(* Logix 5000 project; controller CIP vendor 1 type 14 code 106 rev 20.12; software revision 20.06; part 3 of 13 *)
(* tags used below, declared in another part *)
   Alarm_Preset_Indx : DINT;
   Alarm_Timer : TIMER[128];
   Alarm_Timer_Preset : DINT[128];
   Bit : BOOL[128];
   Counter : COUNTER[10];
   Integer_1 : ALIAS FOR Integer[1];
   Integer_6 : ALIAS FOR Integer[6];
   One_Shot : BOOL[128];
   Panelview : INT[40];
   PV_Current_Select_Step_Op : DINT;
   PV_Edit_Opcodes : DINT[300];
   PV_Edit_Recipe_Name : STRING;
   PV_Edit_Recipe_Top_Row : DINT;
   PV_Edit_Recipes : DINT[7];
   PV_Edit_Recipes_0 : ALIAS FOR PV_Edit_Recipes[0];
   PV_Edit_Recipes_0_Prev : DINT;
   PV_Edit_Screen_Opcodes : DINT[17];
   PV_Edit_Setpoints : REAL[97];
   PV_Edit_Times : DINT[300];
   PV_Rename_Recipe_Name : STRING;
   PV_Security : Security_Main_HMI;
   PV_Security1 : Security_Remote_HMI;
   PV_Step_Time : REAL;
   PV_Visibility : INT[5];
   Recipe : RECIPE[41];
   Recipe_Name : STRING[41];
   Recipe_Name_Indx : DINT;
   SecurityLevel : DINT;
   SecurityLevel1 : DINT;
   Time_Date : DINT[20];
   WashChamberDoorGasketCTRL : DINT;
(* MainProgram, continued *)

ROUTINE _03_PV_SECURITY_REMOTE1_HMI   (* ladder *)
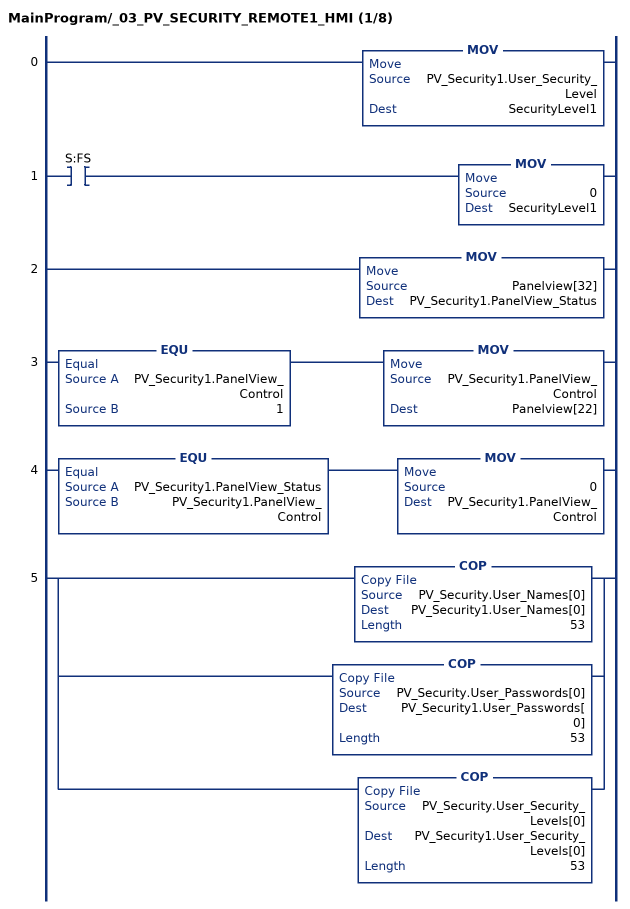
   0: MOV(PV_Security1.User_Security_Level,SecurityLevel1);
   1: XIC(S:FS)MOV(0,SecurityLevel1);
   2: MOV(Panelview[32],PV_Security1.PanelView_Status);
   3: EQU(PV_Security1.PanelView_Control,1)MOV(PV_Security1.PanelView_Control,Panelview[22]);
   4: EQU(PV_Security1.PanelView_Status,PV_Security1.PanelView_Control)MOV(0,PV_Security1.PanelView_Control);
   5: [COP(PV_Security.User_Names[0],PV_Security1.User_Names[0],53) ,COP(PV_Security.User_Passwords[0],PV_Security1.User_Passwords[0],53) ,COP(PV_Security.User_Security_Levels[0],PV_Security1.User_Security_Levels[0],53) ];
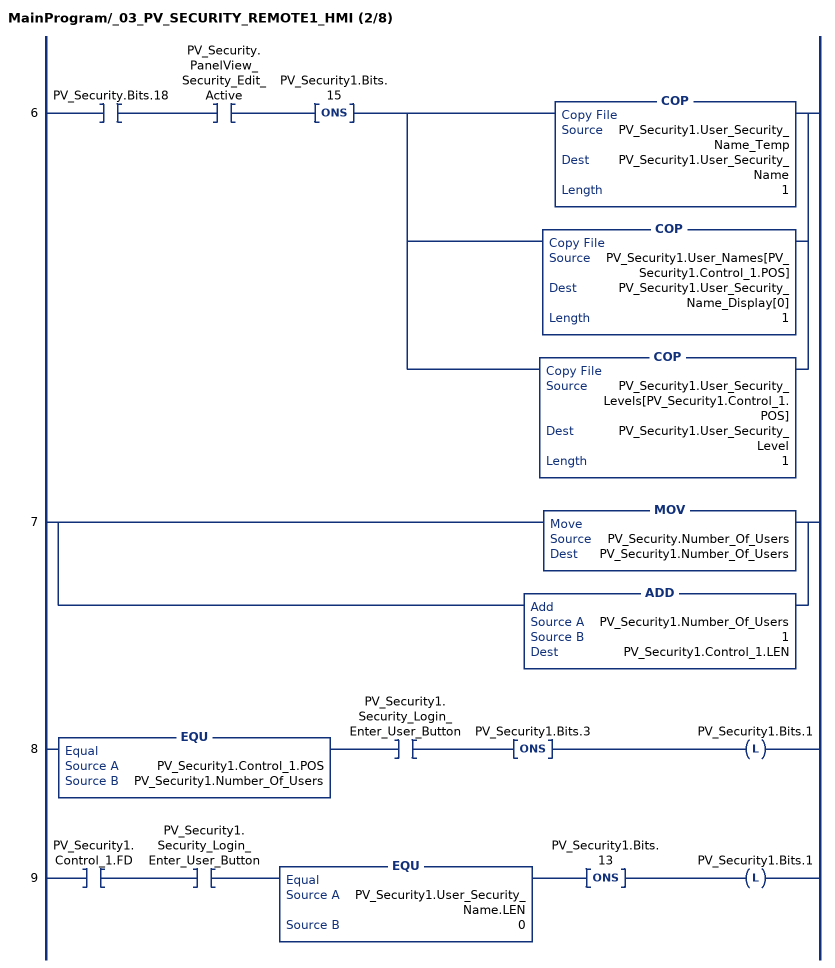
   6: XIC(PV_Security.Bits.18)XIC(PV_Security.PanelView_Security_Edit_Active)ONS(PV_Security1.Bits.15)[COP(PV_Security1.User_Security_Name_Temp,PV_Security1.User_Security_Name,1) ,COP(PV_Security1.User_Names[PV_Security1.Control_1.POS],PV_Security1.User_Security_Name_Display[0],1) ,COP(PV_Security1.User_Security_Levels[PV_Security1.Control_1.POS],PV_Security1.User_Security_Level,1) ];
   7: [MOV(PV_Security.Number_Of_Users,PV_Security1.Number_Of_Users) ,ADD(PV_Security1.Number_Of_Users,1,PV_Security1.Control_1.LEN) ];
   8: EQU(PV_Security1.Control_1.POS,PV_Security1.Number_Of_Users)XIC(PV_Security1.Security_Login_Enter_User_Button)ONS(PV_Security1.Bits.3)OTL(PV_Security1.Bits.1);
   9: XIC(PV_Security1.Control_1.FD)XIC(PV_Security1.Security_Login_Enter_User_Button)EQU(PV_Security1.User_Security_Name.LEN,0)ONS(PV_Security1.Bits.13)OTL(PV_Security1.Bits.1);
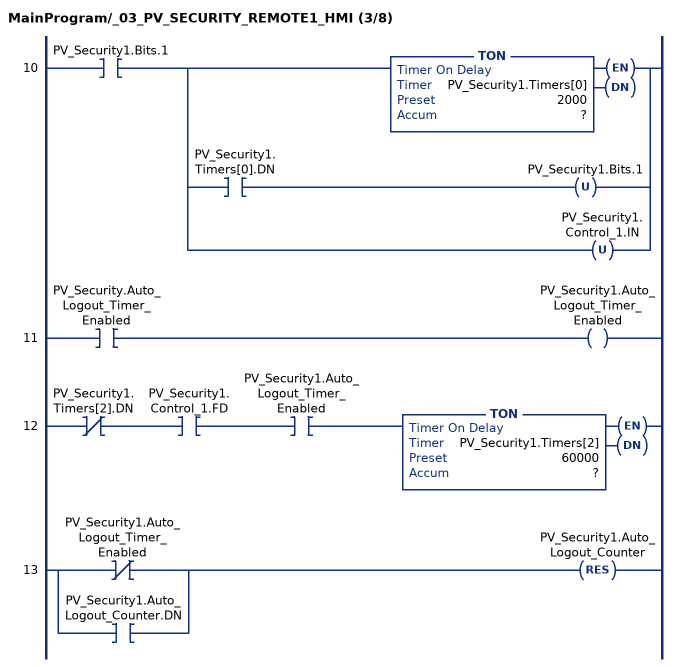
   10: XIC(PV_Security1.Bits.1)[TON(PV_Security1.Timers[0],?,?) ,XIC(PV_Security1.Timers[0].DN) OTU(PV_Security1.Bits.1) ,OTU(PV_Security1.Control_1.IN) ];
   11: XIC(PV_Security.Auto_Logout_Timer_Enabled)OTE(PV_Security1.Auto_Logout_Timer_Enabled);
   12: XIO(PV_Security1.Timers[2].DN)XIC(PV_Security1.Control_1.FD)XIC(PV_Security1.Auto_Logout_Timer_Enabled)TON(PV_Security1.Timers[2],?,?);
   13: [XIO(PV_Security1.Auto_Logout_Timer_Enabled) ,XIC(PV_Security1.Auto_Logout_Counter.DN) ]RES(PV_Security1.Auto_Logout_Counter);
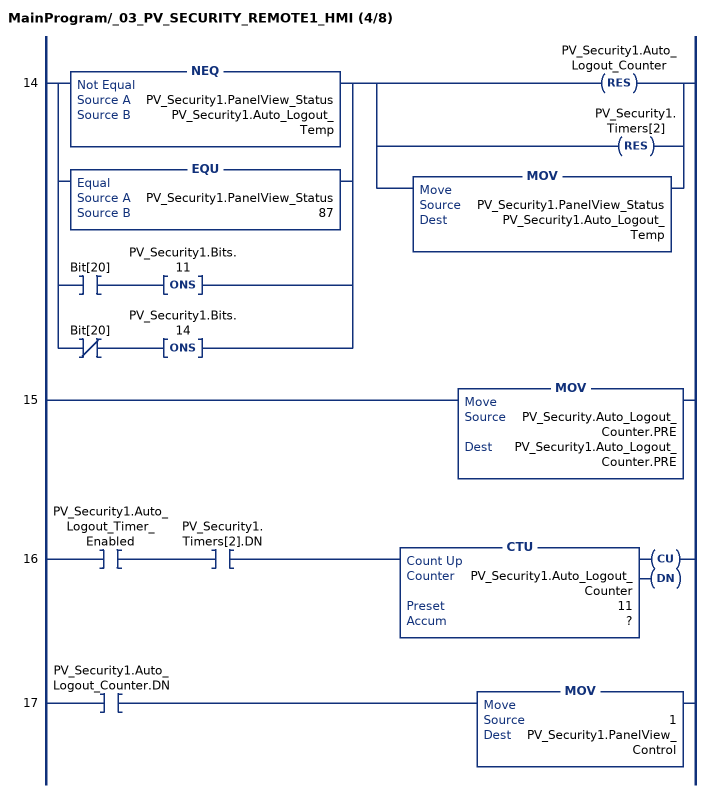
   14: [NEQ(PV_Security1.PanelView_Status,PV_Security1.Auto_Logout_Temp) ,EQU(PV_Security1.PanelView_Status,87) ,XIC(Bit[20]) ONS(PV_Security1.Bits.11) ,XIO(Bit[20]) ONS(PV_Security1.Bits.14) ][RES(PV_Security1.Auto_Logout_Counter) ,RES(PV_Security1.Timers[2]) ,MOV(PV_Security1.PanelView_Status,PV_Security1.Auto_Logout_Temp) ];
   15: MOV(PV_Security.Auto_Logout_Counter.PRE,PV_Security1.Auto_Logout_Counter.PRE);
   16: XIC(PV_Security1.Auto_Logout_Timer_Enabled)XIC(PV_Security1.Timers[2].DN)CTU(PV_Security1.Auto_Logout_Counter,?,?);
   17: XIC(PV_Security1.Auto_Logout_Counter.DN)MOV(1,PV_Security1.PanelView_Control);
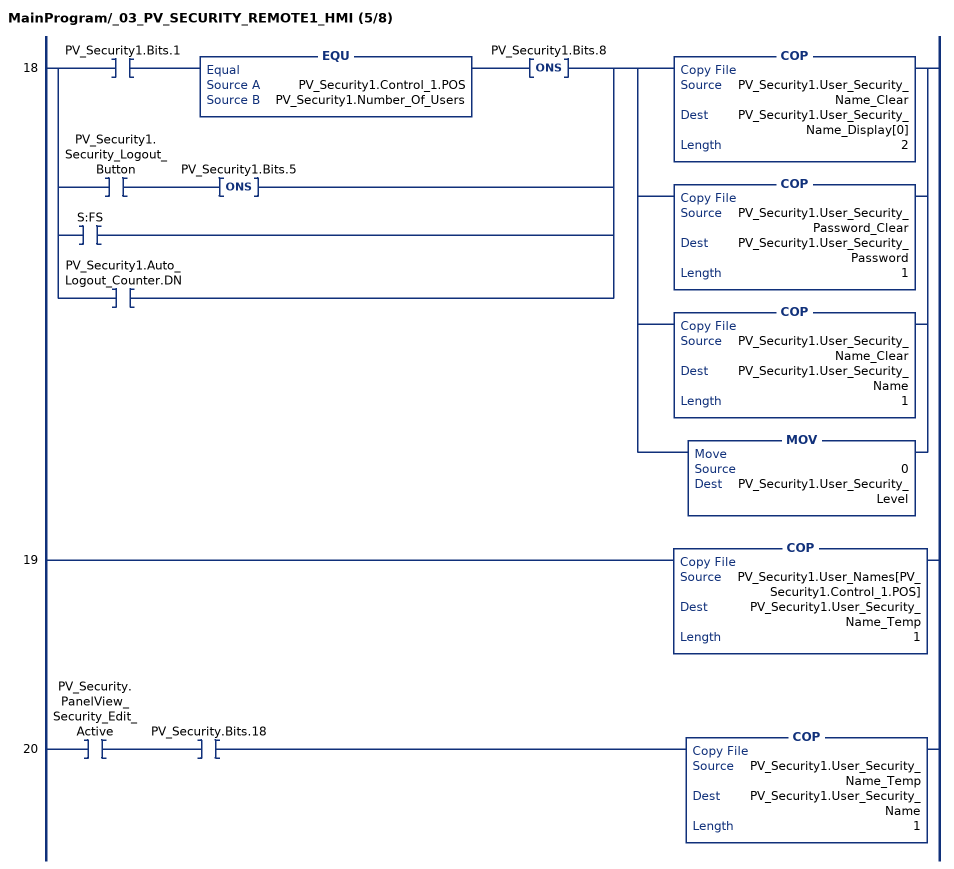
   18: [XIC(PV_Security1.Bits.1) EQU(PV_Security1.Control_1.POS,PV_Security1.Number_Of_Users) ONS(PV_Security1.Bits.8) ,XIC(PV_Security1.Security_Logout_Button) ONS(PV_Security1.Bits.5) ,XIC(S:FS) ,XIC(PV_Security1.Auto_Logout_Counter.DN) ][COP(PV_Security1.User_Security_Name_Clear,PV_Security1.User_Security_Name_Display[0],2) ,COP(PV_Security1.User_Security_Password_Clear,PV_Security1.User_Security_Password,1) ,COP(PV_Security1.User_Security_Name_Clear,PV_Security1.User_Security_Name,1) ,MOV(0,PV_Security1.User_Security_Level) ];
   19: COP(PV_Security1.User_Names[PV_Security1.Control_1.POS],PV_Security1.User_Security_Name_Temp,1);
   20: XIC(PV_Security.PanelView_Security_Edit_Active)XIC(PV_Security.Bits.18)COP(PV_Security1.User_Security_Name_Temp,PV_Security1.User_Security_Name,1);
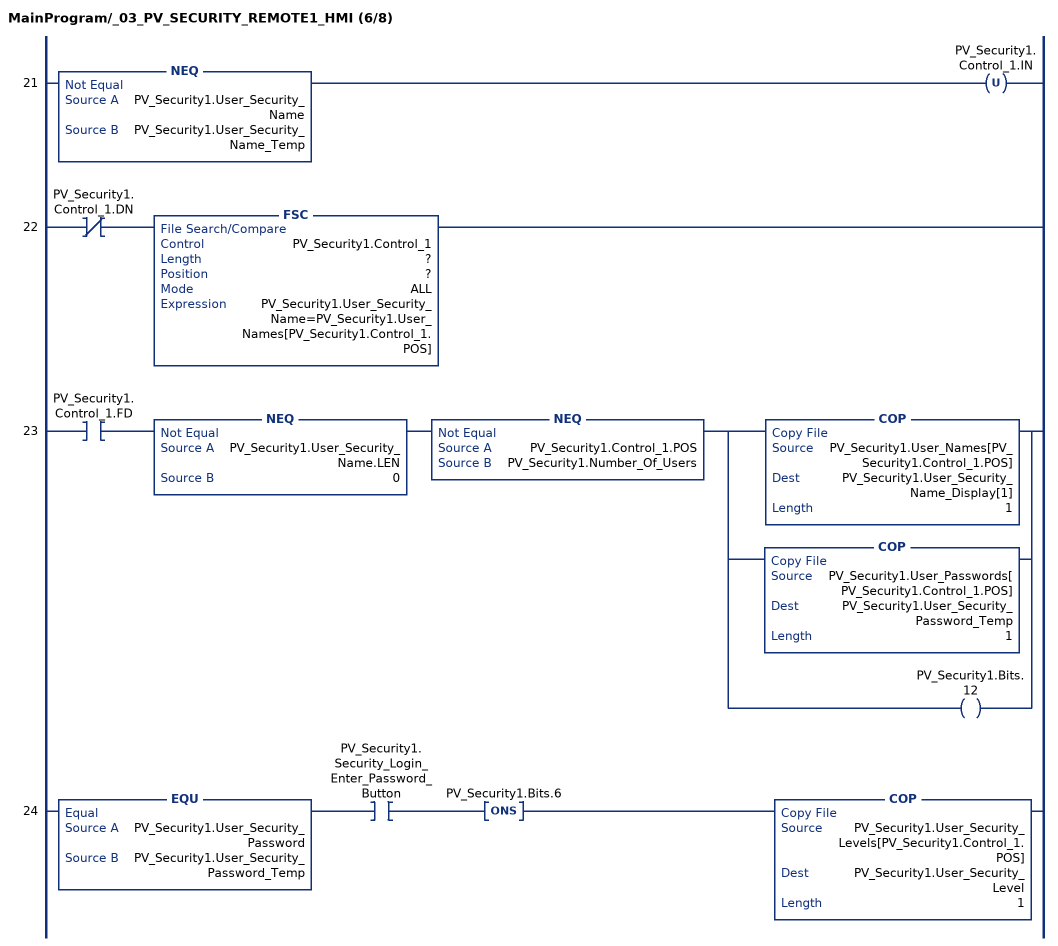
   21: NEQ(PV_Security1.User_Security_Name,PV_Security1.User_Security_Name_Temp)OTU(PV_Security1.Control_1.IN);
   22: XIO(PV_Security1.Control_1.DN)FSC(PV_Security1.Control_1,?,?,ALL,PV_Security1.User_Security_Name=PV_Security1.User_Names[PV_Security1.Control_1.POS]);
   23: XIC(PV_Security1.Control_1.FD)NEQ(PV_Security1.User_Security_Name.LEN,0)NEQ(PV_Security1.Control_1.POS,PV_Security1.Number_Of_Users)[COP(PV_Security1.User_Names[PV_Security1.Control_1.POS],PV_Security1.User_Security_Name_Display[1],1) ,COP(PV_Security1.User_Passwords[PV_Security1.Control_1.POS],PV_Security1.User_Security_Password_Temp,1) ,OTE(PV_Security1.Bits.12) ];
   24: EQU(PV_Security1.User_Security_Password,PV_Security1.User_Security_Password_Temp)XIC(PV_Security1.Security_Login_Enter_Password_Button)ONS(PV_Security1.Bits.6)COP(PV_Security1.User_Security_Levels[PV_Security1.Control_1.POS],PV_Security1.User_Security_Level,1);
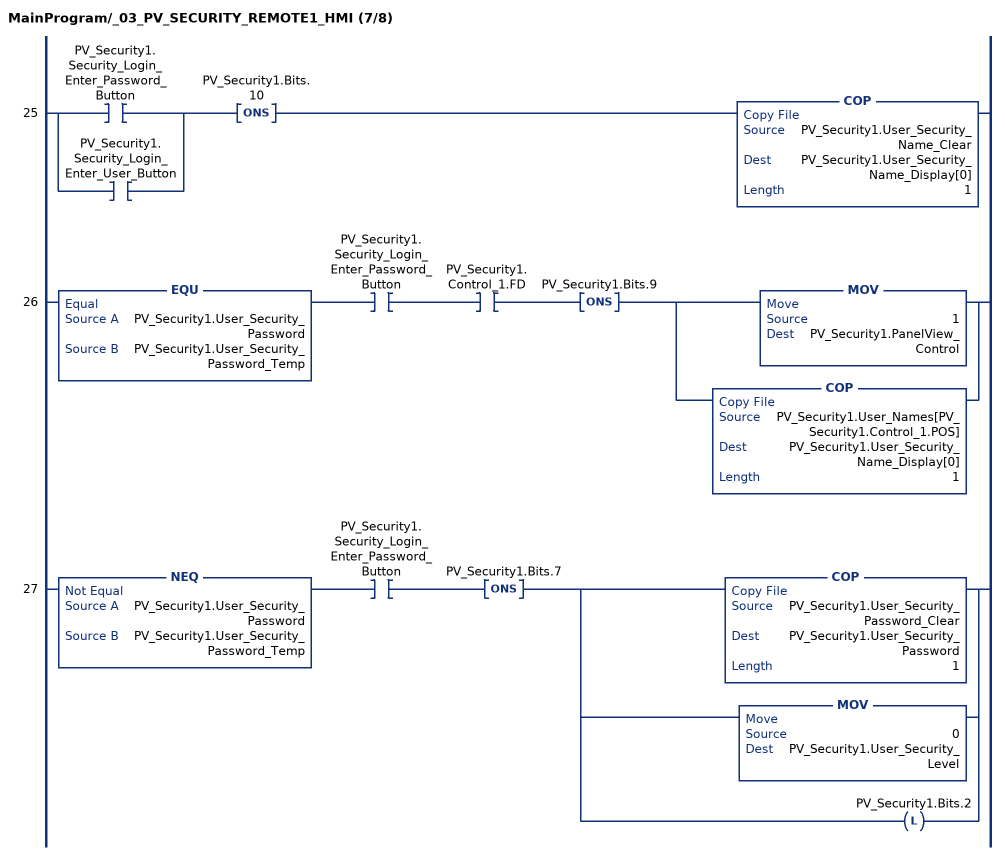
   25: [XIC(PV_Security1.Security_Login_Enter_Password_Button) ,XIC(PV_Security1.Security_Login_Enter_User_Button) ]ONS(PV_Security1.Bits.10)COP(PV_Security1.User_Security_Name_Clear,PV_Security1.User_Security_Name_Display[0],1);
   26: EQU(PV_Security1.User_Security_Password,PV_Security1.User_Security_Password_Temp)XIC(PV_Security1.Security_Login_Enter_Password_Button)XIC(PV_Security1.Control_1.FD)ONS(PV_Security1.Bits.9)[MOV(1,PV_Security1.PanelView_Control) ,COP(PV_Security1.User_Names[PV_Security1.Control_1.POS],PV_Security1.User_Security_Name_Display[0],1) ];
   27: NEQ(PV_Security1.User_Security_Password,PV_Security1.User_Security_Password_Temp)XIC(PV_Security1.Security_Login_Enter_Password_Button)ONS(PV_Security1.Bits.7)[COP(PV_Security1.User_Security_Password_Clear,PV_Security1.User_Security_Password,1) ,MOV(0,PV_Security1.User_Security_Level) ,OTL(PV_Security1.Bits.2) ];
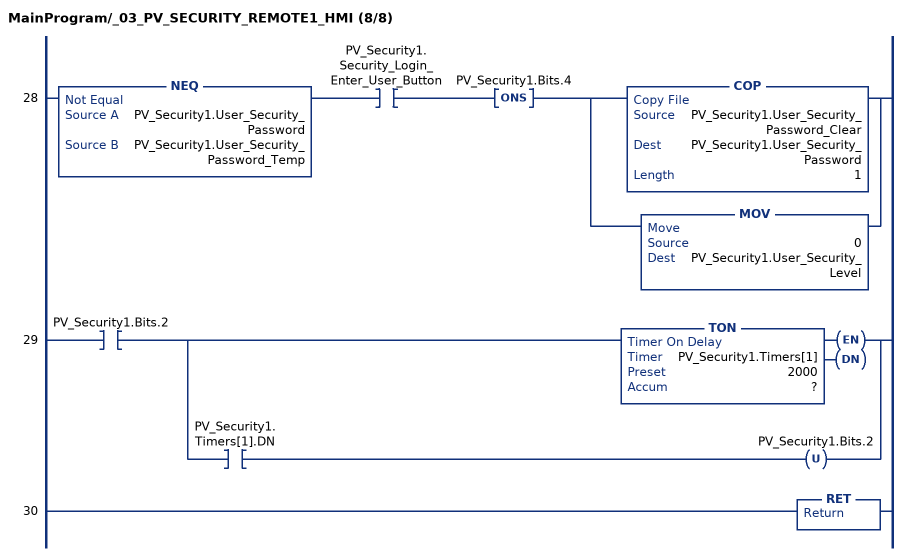
   28: NEQ(PV_Security1.User_Security_Password,PV_Security1.User_Security_Password_Temp)XIC(PV_Security1.Security_Login_Enter_User_Button)ONS(PV_Security1.Bits.4)[COP(PV_Security1.User_Security_Password_Clear,PV_Security1.User_Security_Password,1) ,MOV(0,PV_Security1.User_Security_Level) ];
   29: XIC(PV_Security1.Bits.2)[TON(PV_Security1.Timers[1],?,?) ,XIC(PV_Security1.Timers[1].DN) OTU(PV_Security1.Bits.2) ];
   30: RET();
END_ROUTINE

ROUTINE _04_PVPLUS   (* ladder *)
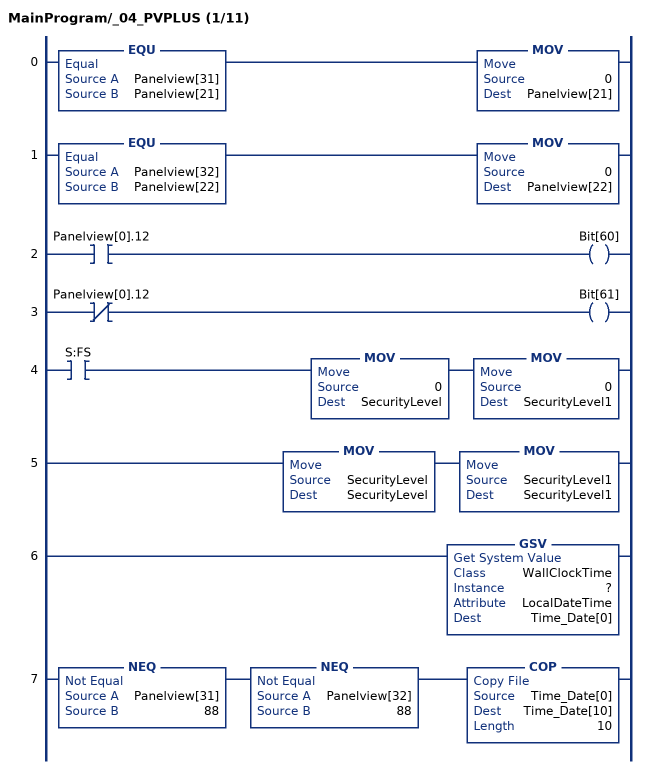
   0: EQU(Panelview[31],Panelview[21])MOV(0,Panelview[21]);
   1: EQU(Panelview[32],Panelview[22])MOV(0,Panelview[22]);
   2: XIC(Panelview[0].12)OTE(Bit[60]);
   3: XIO(Panelview[0].12)OTE(Bit[61]);
   4: XIC(S:FS)MOV(0,SecurityLevel)MOV(0,SecurityLevel1);
   5: MOV(SecurityLevel,SecurityLevel)MOV(SecurityLevel1,SecurityLevel1);
   6: GSV(WallClockTime,?,LocalDateTime,Time_Date[0]);
   7: NEQ(Panelview[31],88)NEQ(Panelview[32],88)COP(Time_Date[0],Time_Date[10],10);
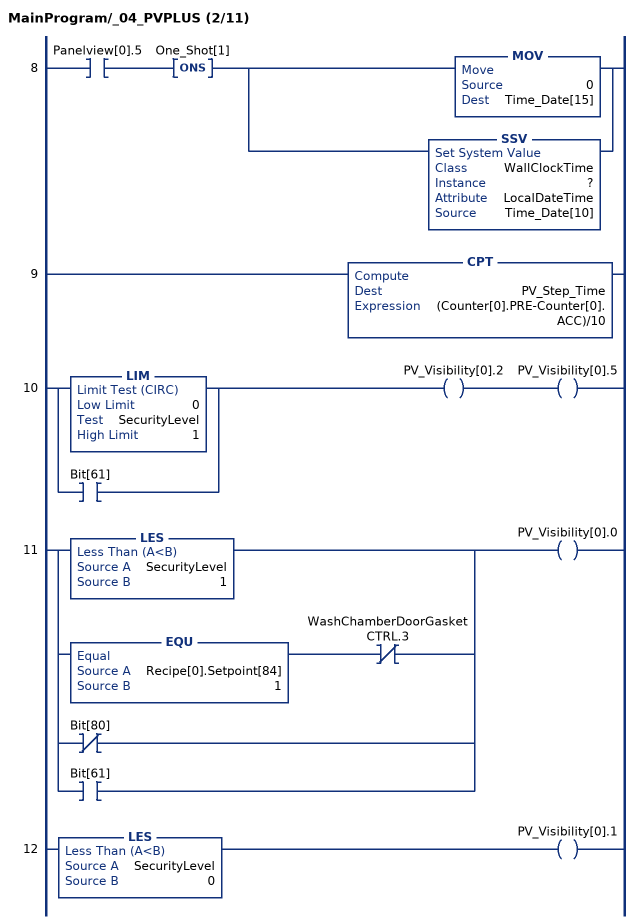
   8: XIC(Panelview[0].5)ONS(One_Shot[1])[MOV(0,Time_Date[15]) ,SSV(WallClockTime,?,LocalDateTime,Time_Date[10]) ];
   9: CPT(PV_Step_Time,(Counter[0].PRE-Counter[0].ACC)/10);
   10: [LIM(0,SecurityLevel,1) ,XIC(Bit[61]) ]OTE(PV_Visibility[0].2)OTE(PV_Visibility[0].5);
   11: [LES(SecurityLevel,1) ,EQU(Recipe[0].Setpoint[84],1) XIO(WashChamberDoorGasketCTRL.3) ,XIO(Bit[80]) ,XIC(Bit[61]) ]OTE(PV_Visibility[0].0);
   12: LES(SecurityLevel,0)OTE(PV_Visibility[0].1);
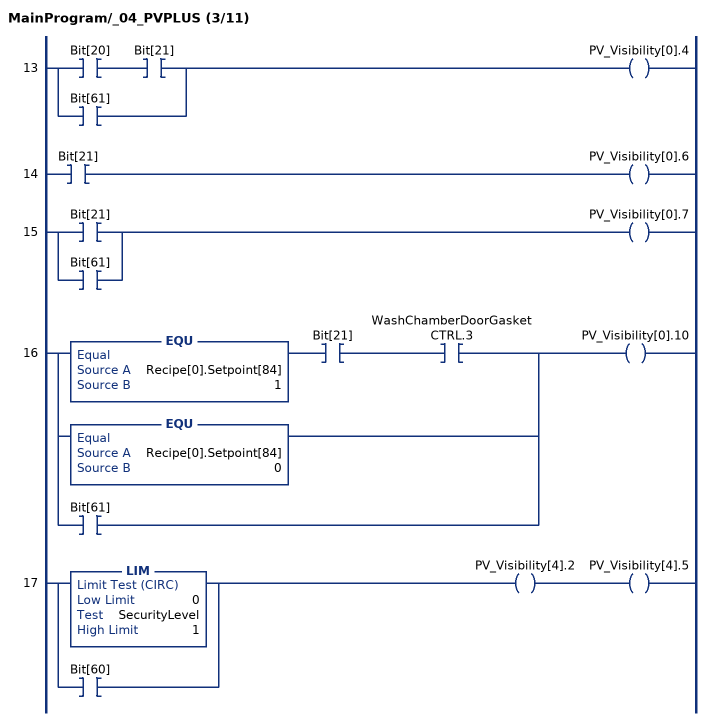
   13: [XIC(Bit[20]) XIC(Bit[21]) ,XIC(Bit[61]) ]OTE(PV_Visibility[0].4);
   14: XIC(Bit[21])OTE(PV_Visibility[0].6);
   15: [XIC(Bit[21]) ,XIC(Bit[61]) ]OTE(PV_Visibility[0].7);
   16: [EQU(Recipe[0].Setpoint[84],1) XIC(Bit[21]) XIC(WashChamberDoorGasketCTRL.3) ,EQU(Recipe[0].Setpoint[84],0) ,XIC(Bit[61]) ]OTE(PV_Visibility[0].10);
   17: [LIM(0,SecurityLevel,1) ,XIC(Bit[60]) ]OTE(PV_Visibility[4].2)OTE(PV_Visibility[4].5);
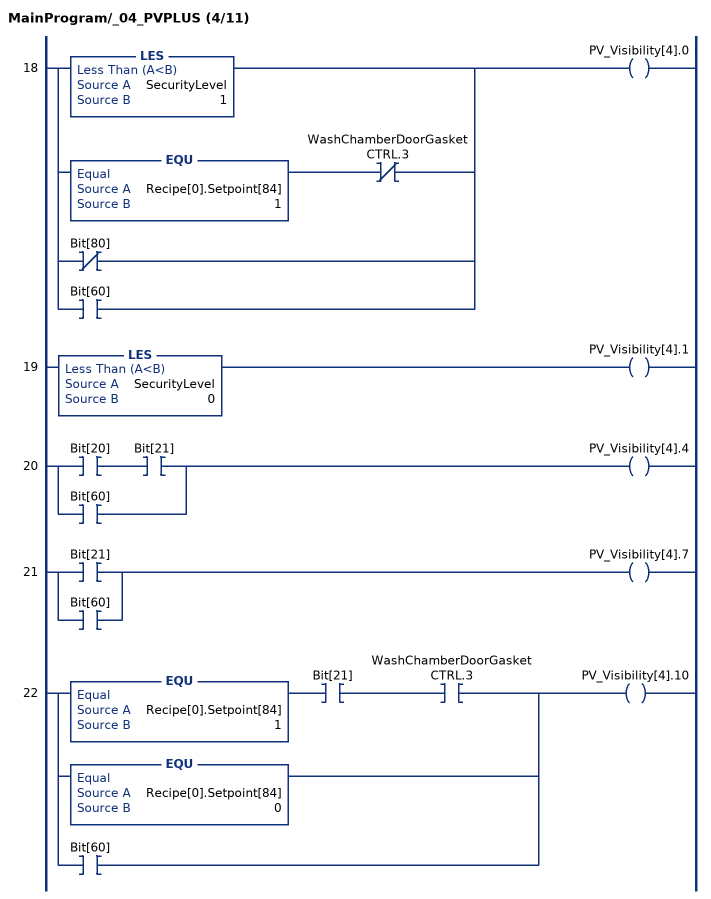
   18: [LES(SecurityLevel,1) ,EQU(Recipe[0].Setpoint[84],1) XIO(WashChamberDoorGasketCTRL.3) ,XIO(Bit[80]) ,XIC(Bit[60]) ]OTE(PV_Visibility[4].0);
   19: LES(SecurityLevel,0)OTE(PV_Visibility[4].1);
   20: [XIC(Bit[20]) XIC(Bit[21]) ,XIC(Bit[60]) ]OTE(PV_Visibility[4].4);
   21: [XIC(Bit[21]) ,XIC(Bit[60]) ]OTE(PV_Visibility[4].7);
   22: [EQU(Recipe[0].Setpoint[84],1) XIC(Bit[21]) XIC(WashChamberDoorGasketCTRL.3) ,EQU(Recipe[0].Setpoint[84],0) ,XIC(Bit[60]) ]OTE(PV_Visibility[4].10);
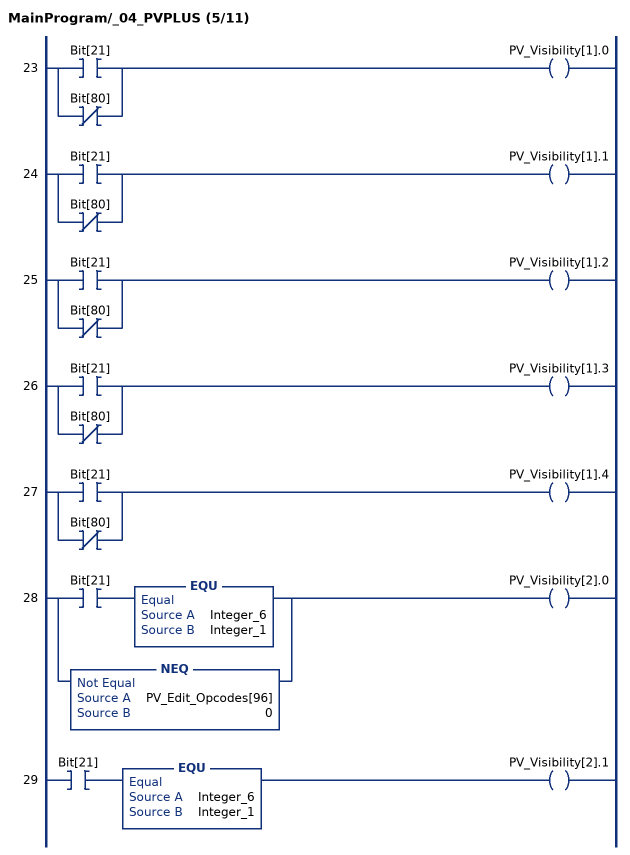
   23: [XIC(Bit[21]) ,XIO(Bit[80]) ]OTE(PV_Visibility[1].0);
   24: [XIC(Bit[21]) ,XIO(Bit[80]) ]OTE(PV_Visibility[1].1);
   25: [XIC(Bit[21]) ,XIO(Bit[80]) ]OTE(PV_Visibility[1].2);
   26: [XIC(Bit[21]) ,XIO(Bit[80]) ]OTE(PV_Visibility[1].3);
   27: [XIC(Bit[21]) ,XIO(Bit[80]) ]OTE(PV_Visibility[1].4);
   28: [XIC(Bit[21]) EQU(Integer_6,Integer_1) ,NEQ(PV_Edit_Opcodes[96],0) ]OTE(PV_Visibility[2].0);
   29: XIC(Bit[21])EQU(Integer_6,Integer_1)OTE(PV_Visibility[2].1);
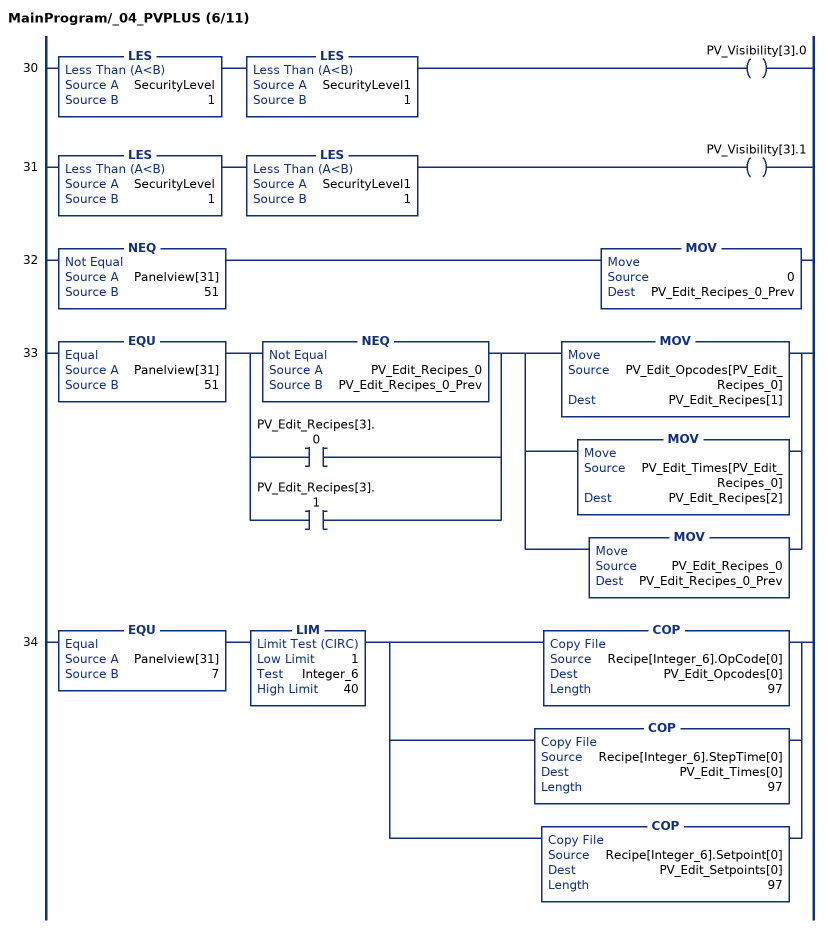
   30: LES(SecurityLevel,1)LES(SecurityLevel1,1)OTE(PV_Visibility[3].0);
   31: LES(SecurityLevel,1)LES(SecurityLevel1,1)OTE(PV_Visibility[3].1);
   32: NEQ(Panelview[31],51)MOV(0,PV_Edit_Recipes_0_Prev);
   33: EQU(Panelview[31],51)[NEQ(PV_Edit_Recipes_0,PV_Edit_Recipes_0_Prev) ,XIC(PV_Edit_Recipes[3].0) ,XIC(PV_Edit_Recipes[3].1) ][MOV(PV_Edit_Opcodes[PV_Edit_Recipes_0],PV_Edit_Recipes[1]) ,MOV(PV_Edit_Times[PV_Edit_Recipes_0],PV_Edit_Recipes[2]) ,MOV(PV_Edit_Recipes_0,PV_Edit_Recipes_0_Prev) ];
   34: EQU(Panelview[31],7)LIM(1,Integer_6,40)[COP(Recipe[Integer_6].OpCode[0],PV_Edit_Opcodes[0],97) ,COP(Recipe[Integer_6].StepTime[0],PV_Edit_Times[0],97) ,COP(Recipe[Integer_6].Setpoint[0],PV_Edit_Setpoints[0],97) ];
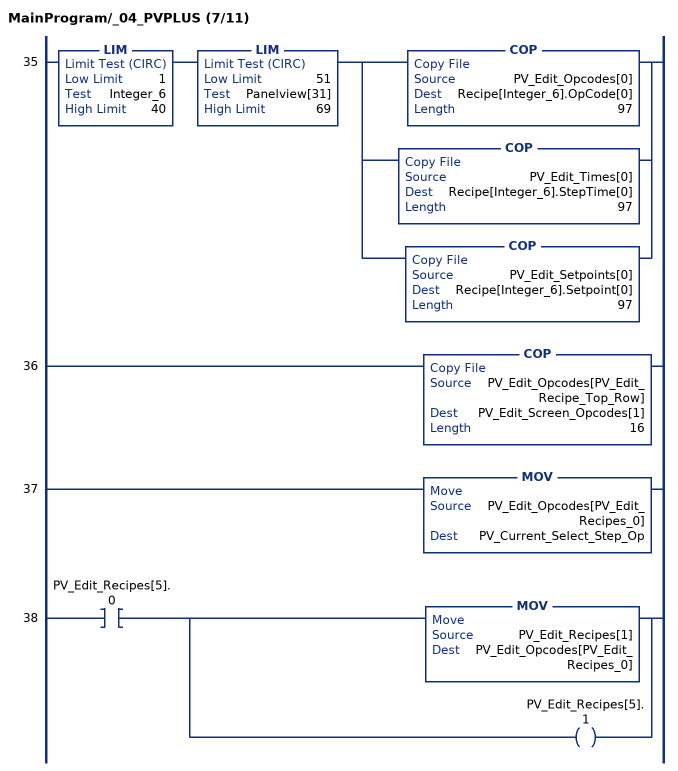
   35: LIM(1,Integer_6,40)LIM(51,Panelview[31],69)[COP(PV_Edit_Opcodes[0],Recipe[Integer_6].OpCode[0],97) ,COP(PV_Edit_Times[0],Recipe[Integer_6].StepTime[0],97) ,COP(PV_Edit_Setpoints[0],Recipe[Integer_6].Setpoint[0],97) ];
   36: COP(PV_Edit_Opcodes[PV_Edit_Recipe_Top_Row],PV_Edit_Screen_Opcodes[1],16);
   37: MOV(PV_Edit_Opcodes[PV_Edit_Recipes_0],PV_Current_Select_Step_Op);
   38: XIC(PV_Edit_Recipes[5].0)[MOV(PV_Edit_Recipes[1],PV_Edit_Opcodes[PV_Edit_Recipes_0]) ,OTE(PV_Edit_Recipes[5].1) ];
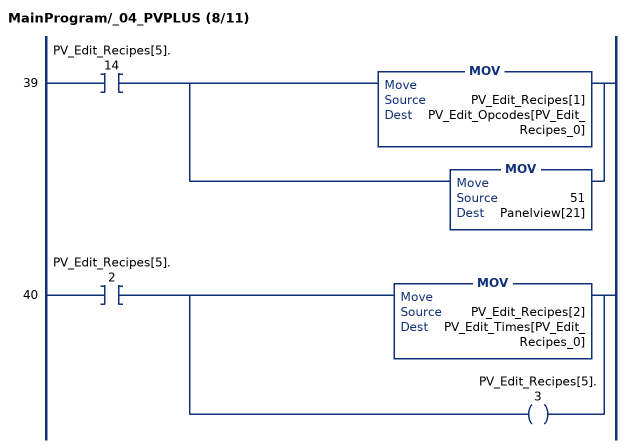
   39: XIC(PV_Edit_Recipes[5].14)[MOV(PV_Edit_Recipes[1],PV_Edit_Opcodes[PV_Edit_Recipes_0]) ,MOV(51,Panelview[21]) ];
   40: XIC(PV_Edit_Recipes[5].2)[MOV(PV_Edit_Recipes[2],PV_Edit_Times[PV_Edit_Recipes_0]) ,OTE(PV_Edit_Recipes[5].3) ];
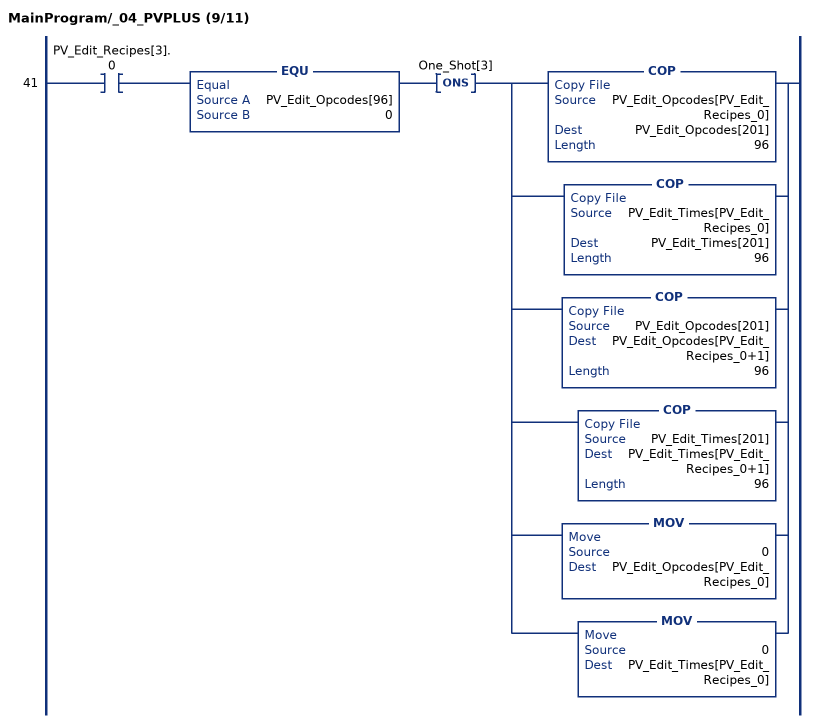
   41: XIC(PV_Edit_Recipes[3].0)EQU(PV_Edit_Opcodes[96],0)ONS(One_Shot[3])[COP(PV_Edit_Opcodes[PV_Edit_Recipes_0],PV_Edit_Opcodes[201],96) ,COP(PV_Edit_Times[PV_Edit_Recipes_0],PV_Edit_Times[201],96) ,COP(PV_Edit_Opcodes[201],PV_Edit_Opcodes[PV_Edit_Recipes_0+1],96) ,COP(PV_Edit_Times[201],PV_Edit_Times[PV_Edit_Recipes_0+1],96) ,MOV(0,PV_Edit_Opcodes[PV_Edit_Recipes_0]) ,MOV(0,PV_Edit_Times[PV_Edit_Recipes_0]) ];
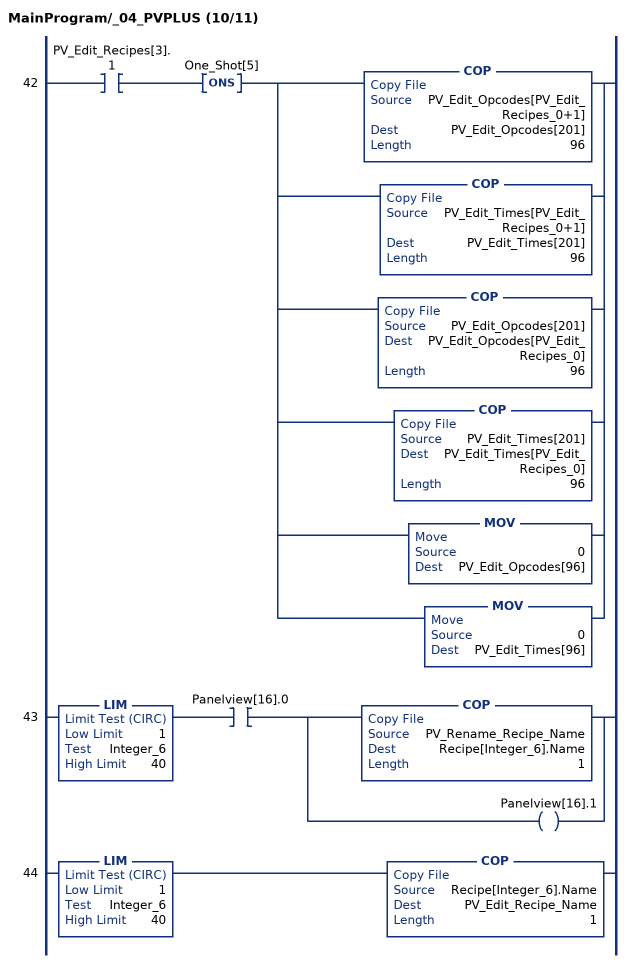
   42: XIC(PV_Edit_Recipes[3].1)ONS(One_Shot[5])[COP(PV_Edit_Opcodes[PV_Edit_Recipes_0+1],PV_Edit_Opcodes[201],96) ,COP(PV_Edit_Times[PV_Edit_Recipes_0+1],PV_Edit_Times[201],96) ,COP(PV_Edit_Opcodes[201],PV_Edit_Opcodes[PV_Edit_Recipes_0],96) ,COP(PV_Edit_Times[201],PV_Edit_Times[PV_Edit_Recipes_0],96) ,MOV(0,PV_Edit_Opcodes[96]) ,MOV(0,PV_Edit_Times[96]) ];
   43: LIM(1,Integer_6,40)XIC(Panelview[16].0)[COP(PV_Rename_Recipe_Name,Recipe[Integer_6].Name,1) ,OTE(Panelview[16].1) ];
   44: LIM(1,Integer_6,40)COP(Recipe[Integer_6].Name,PV_Edit_Recipe_Name,1);
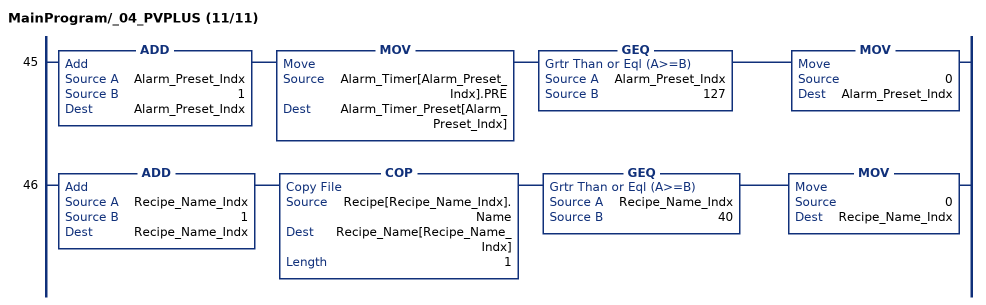
   45: ADD(Alarm_Preset_Indx,1,Alarm_Preset_Indx)MOV(Alarm_Timer[Alarm_Preset_Indx].PRE,Alarm_Timer_Preset[Alarm_Preset_Indx])GEQ(Alarm_Preset_Indx,127)MOV(0,Alarm_Preset_Indx);
   46: ADD(Recipe_Name_Indx,1,Recipe_Name_Indx)COP(Recipe[Recipe_Name_Indx].Name,Recipe_Name[Recipe_Name_Indx],1)GEQ(Recipe_Name_Indx,40)MOV(0,Recipe_Name_Indx);
END_ROUTINE
